(* IEC 61131-3 sources: codesys-api/examples/plc_architecture/bench/st, 5 files *)

(* ---- PRG_BusTask.st ---- *)
PROGRAM PRG_BusTask
// Body of the bus task on the bench (BusTask: cyclic 5 ms, priority between control and comms): PRG_Bus, timed.
// ExecUs is wall time, so it includes time the control task preempted it. Per line: requests and errors per
// second over the last full second, and how long the slowest request took.
VAR
	ResetStats : BOOL;
	ScanCount : UDINT;
	ExecUs : UDINT;
	MaxExecUs : UDINT;
	ExecTotalUs : ULINT;
	MaxIntervalUs : UDINT;
	RequestsPerSecond : ARRAY[1..GVL_Bus.LINE_COUNT] OF UDINT;
	ErrorsPerSecond : ARRAY[1..GVL_Bus.LINE_COUNT] OF UDINT;

	StartUs : ULINT;
	PreviousStartUs : ULINT;
	SecondStartUs : ULINT;
	RequestsAtSecond : ARRAY[1..GVL_Bus.LINE_COUNT] OF UDINT;
	ErrorsAtSecond : ARRAY[1..GVL_Bus.LINE_COUNT] OF UDINT;
	Index : INT;
END_VAR
// ---- implementation ----
StartUs := F_NowUs();
IF ResetStats THEN
	ResetStats := FALSE;
	ScanCount := 0;
	MaxExecUs := 0;
	ExecTotalUs := 0;
	MaxIntervalUs := 0;
	PreviousStartUs := 0;
END_IF
IF PreviousStartUs <> 0 THEN
	MaxIntervalUs := MAX(MaxIntervalUs, ULINT_TO_UDINT(StartUs - PreviousStartUs));
END_IF
PreviousStartUs := StartUs;

PRG_Bus();
PRG_SerialProbe();       // idle unless IsEnabled

IF StartUs - SecondStartUs >= 1000000 THEN
	SecondStartUs := StartUs;
	FOR Index := 1 TO GVL_Bus.LINE_COUNT DO
		RequestsPerSecond[Index] := PRG_Bus.Lines[Index].RequestCount - RequestsAtSecond[Index];
		ErrorsPerSecond[Index] := PRG_Bus.Lines[Index].ErrorCount - ErrorsAtSecond[Index];
		RequestsAtSecond[Index] := PRG_Bus.Lines[Index].RequestCount;
		ErrorsAtSecond[Index] := PRG_Bus.Lines[Index].ErrorCount;
	END_FOR
END_IF

ExecUs := ULINT_TO_UDINT(F_NowUs() - StartUs);
MaxExecUs := MAX(MaxExecUs, ExecUs);
ExecTotalUs := ExecTotalUs + ExecUs;
ScanCount := ScanCount + 1;

(* ---- PRG_CommsTask.st ---- *)
PROGRAM PRG_CommsTask
// Body of the comms task on the two-task bench (CommsTask: cyclic, priority below the control task):
// PRG_Comms, timed. ExecUs is wall time from start to end of this task's scan, so it includes any time the
// control task preempted it. A publish is timed from PRG_Comms.IsRequested going TRUE to FALSE (done).
VAR
	IsEnabled : BOOL := TRUE;
	ResetStats : BOOL;

	ScanCount : UDINT;
	ExecUs : UDINT;
	MaxExecUs : UDINT;
	ExecTotalUs : ULINT;
	MaxIntervalUs : UDINT;
	PublishCount : UDINT;
	LastPublishUs : UDINT;
	MaxPublishUs : UDINT;
	LastPayloadLength : UDINT;
	MaxClientCalls : INT;

	StartUs : ULINT;
	PreviousStartUs : ULINT;
	RequestUs : ULINT;
	WasRequested : BOOL;
END_VAR
// ---- implementation ----
StartUs := F_NowUs();
IF ResetStats THEN
	ResetStats := FALSE;
	ScanCount := 0;
	MaxExecUs := 0;
	ExecTotalUs := 0;
	MaxIntervalUs := 0;
	PublishCount := 0;
	MaxPublishUs := 0;
	MaxClientCalls := 0;
	PreviousStartUs := 0;
END_IF
IF PreviousStartUs <> 0 THEN
	MaxIntervalUs := MAX(MaxIntervalUs, ULINT_TO_UDINT(StartUs - PreviousStartUs));
END_IF
PreviousStartUs := StartUs;

IF IsEnabled THEN
	PRG_Comms();
	MaxClientCalls := MAX(MaxClientCalls, PRG_Comms.ClientCall);
	IF PRG_Comms.IsRequested AND NOT WasRequested THEN
		RequestUs := StartUs;
		LastPayloadLength := PRG_Comms.Used;
	ELSIF WasRequested AND NOT PRG_Comms.IsRequested THEN
		LastPublishUs := ULINT_TO_UDINT(StartUs - RequestUs);
		MaxPublishUs := MAX(MaxPublishUs, LastPublishUs);
		PublishCount := PublishCount + 1;
	END_IF
	WasRequested := PRG_Comms.IsRequested;
END_IF

ExecUs := ULINT_TO_UDINT(F_NowUs() - StartUs);
MaxExecUs := MAX(MaxExecUs, ExecUs);
ExecTotalUs := ExecTotalUs + ExecUs;
ScanCount := ScanCount + 1;

(* ---- PRG_ControlTask.st ---- *)
PROGRAM PRG_ControlTask
// Body of the control task on the two-task bench (MainTask: cyclic 50 ms, priority 1): simulated inputs,
// then the control pipeline, timed. IntervalUs is the start-to-start time of this task; its deviation from
// NominalUs is the jitter the comms task could cause. ExecUs is the time spent in the task.
VAR
	NominalUs : ULINT := 50000;         // the task's configured interval
	ResetStats : BOOL;
	IsQualityCountRequested : BOOL;     // count tags per quality once (costs a pass over the table)

	ScanCount : UDINT;
	IntervalUs : UDINT;
	MinIntervalUs : UDINT := 16#FFFFFFFF;
	MaxIntervalUs : UDINT;
	MaxDeviationUs : UDINT;             // largest |IntervalUs - NominalUs|
	// |IntervalUs - NominalUs| in bands: <= 0.1 ms, 0.5 ms, 1 ms, 2 ms, 5 ms, more
	Deviation : ARRAY[0..5] OF UDINT;
	ExecUs : UDINT;
	MaxExecUs : UDINT;
	ExecTotalUs : ULINT;
	SimUs : UDINT;
	MaxSimUs : UDINT;
	GoodCount : INT;
	NotGoodCount : INT;

	StartUs : ULINT;
	PreviousStartUs : ULINT;
	StepUs : ULINT;
	DeviationUs : UDINT;
	Index : INT;
END_VAR
// ---- implementation ----
StartUs := F_NowUs();
IF ResetStats THEN
	ResetStats := FALSE;
	ScanCount := 0;
	MinIntervalUs := 16#FFFFFFFF;
	MaxIntervalUs := 0;
	MaxDeviationUs := 0;
	FOR Index := 0 TO 5 DO
		Deviation[Index] := 0;
	END_FOR
	MaxExecUs := 0;
	ExecTotalUs := 0;
	MaxSimUs := 0;
	PreviousStartUs := 0;
END_IF
IF PreviousStartUs <> 0 THEN
	IntervalUs := ULINT_TO_UDINT(StartUs - PreviousStartUs);
	MinIntervalUs := MIN(MinIntervalUs, IntervalUs);
	MaxIntervalUs := MAX(MaxIntervalUs, IntervalUs);
	IF UDINT_TO_ULINT(IntervalUs) >= NominalUs THEN
		DeviationUs := IntervalUs - ULINT_TO_UDINT(NominalUs);
	ELSE
		DeviationUs := ULINT_TO_UDINT(NominalUs) - IntervalUs;
	END_IF
	MaxDeviationUs := MAX(MaxDeviationUs, DeviationUs);
	IF DeviationUs <= 100 THEN
		Deviation[0] := Deviation[0] + 1;
	ELSIF DeviationUs <= 500 THEN
		Deviation[1] := Deviation[1] + 1;
	ELSIF DeviationUs <= 1000 THEN
		Deviation[2] := Deviation[2] + 1;
	ELSIF DeviationUs <= 2000 THEN
		Deviation[3] := Deviation[3] + 1;
	ELSIF DeviationUs <= 5000 THEN
		Deviation[4] := Deviation[4] + 1;
	ELSE
		Deviation[5] := Deviation[5] + 1;
	END_IF
END_IF
PreviousStartUs := StartUs;

StepUs := F_NowUs();
PRG_SimInputs();
SimUs := ULINT_TO_UDINT(F_NowUs() - StepUs);
MaxSimUs := MAX(MaxSimUs, SimUs);

PRG_Control();

IF IsQualityCountRequested THEN
	IsQualityCountRequested := FALSE;
	GoodCount := 0;
	NotGoodCount := 0;
	FOR Index := 1 TO GVL_Tags.TAG_COUNT DO
		IF GVL_Tags.Tags[Index].Quality = E_Quality.GOOD THEN
			GoodCount := GoodCount + 1;
		ELSE
			NotGoodCount := NotGoodCount + 1;
		END_IF
	END_FOR
END_IF

ExecUs := ULINT_TO_UDINT(F_NowUs() - StartUs);
MaxExecUs := MAX(MaxExecUs, ExecUs);
ExecTotalUs := ExecTotalUs + ExecUs;
ScanCount := ScanCount + 1;

(* ---- PRG_SerialProbe.st ---- *)
PROGRAM PRG_SerialProbe
// Receive-only check of a PLC serial port, no Modbus: opens the port with SysCom and counts every byte that
// arrives, keeping the last 32. For "the PLC sends but never hears a reply": send a known pattern from the PC
// (bench/serial_pattern.py) and see whether it lands here. Turn the bus line on that port off first
// (PRG_Bus.Lines[n].IsEnabled := FALSE); a port can only be open once. Called from the bus task.
VAR
	IsEnabled : BOOL;                   // set online
	ComPort : INT := 2;
	Baudrate : UDINT := 9600;
	IsVendorSequence : BOOL := TRUE;    // open like AutomationDirect's example (SysComOpen + SysComSetSettings)
	SetResult : UDINT;

	IsOpen : BOOL;
	OpenResult : UDINT;                 // runtime error code of the last open; 0 = OK
	BytesReceived : UDINT;
	ReadCalls : UDINT;
	LastBytes : ARRAY[0..31] OF BYTE;   // most recent bytes, oldest overwritten first
	NextSlot : INT;

	Handle : SysCom.RTS_IEC_HANDLE;
	Settings : SysCom.SysComSettings;
	Result : SysCom.RTS_IEC_RESULT;
	Buffer : ARRAY[0..63] OF BYTE;
	Count : UDINT;
	Index : UDINT;
END_VAR
// ---- implementation ----
IF IsEnabled AND NOT IsOpen THEN
	Settings.sPort := SysCom.SYS_COM_PORTS.SYS_COMPORT1;
	IF ComPort = 2 THEN
		Settings.sPort := SysCom.SYS_COM_PORTS.SYS_COMPORT2;
	END_IF
	Settings.ulBaudrate := SysCom.SYS_COM_BAUDRATE.SYS_BR_9600;
	IF Baudrate = 115200 THEN
		Settings.ulBaudrate := SysCom.SYS_COM_BAUDRATE.SYS_BR_115200;
	END_IF
	Settings.byParity := SysCom.SYS_COM_PARITY.SYS_NOPARITY;
	Settings.byStopBits := SysCom.SYS_COM_STOPBITS.SYS_ONESTOPBIT;
	Settings.ulTimeout := 0;
	Settings.ulBufferSize := 0;
	IF IsVendorSequence THEN
		// AutomationDirect's Demo_SerialPassthrough: open the port, then apply the settings.
		Settings.ulTimeout := 10;
		Handle := SysCom.SysComOpen(sPort := Settings.sPort, pResult := ADR(Result));
		OpenResult := Result;
		IF Result = 0 THEN
			Result := SysCom.SysComSetSettings(hCom := Handle, pSettings := ADR(Settings), pSettingsEx := 0);
			SetResult := Result;
		END_IF
	ELSE
		Handle := SysCom.SysComOpen2(pSettings := ADR(Settings), pSettingsEx := 0, pResult := ADR(Result));
		OpenResult := Result;
	END_IF
	IsOpen := Result = 0;
ELSIF NOT IsEnabled AND IsOpen THEN
	SysCom.SysComClose(hCom := Handle);
	IsOpen := FALSE;
END_IF

IF IsOpen THEN
	Count := SysCom.SysComRead(hCom := Handle, pbyBuffer := ADR(Buffer), ulSize := SIZEOF(Buffer), ulTimeout := 0, pResult := ADR(Result));
	ReadCalls := ReadCalls + 1;
	IF Count > 0 THEN
		FOR Index := 0 TO MIN(Count, SIZEOF(Buffer)) - 1 DO
			LastBytes[NextSlot] := Buffer[Index];
			NextSlot := (NextSlot + 1) MOD 32;
		END_FOR
		BytesReceived := BytesReceived + Count;
	END_IF
END_IF

(* ---- PRG_SimInputs.st ---- *)
PROGRAM PRG_SimInputs
// Bench stand-in for local I/O: the tags of source 0 keep moving. Each scan ChangePerScan of them get a new raw
// value, cycling through the table (100 per 50 ms scan = every tag changes about once a second). Tags of the bus
// devices come from PRG_Bus instead. Values stay inside the generated ranges: BOOL 0/1, INT 0..99,999, REAL raw
// 0..4,999 (scale 0.1 -> 0..499.9).
VAR
	ChangePerScan : INT := 100;
	NextIndex : INT := 1;
	Step : DINT;
	Count : INT;
END_VAR
// ---- implementation ----
Step := Step + 1;
FOR Count := 1 TO ChangePerScan DO
	IF GVL_Tags.TagConfig[NextIndex].Source = 0 THEN
		CASE GVL_Tags.TagConfig[NextIndex].Kind OF
			E_TagKind.BOOL_TAG:
				GVL_Tags.RawInputs[NextIndex] := DINT_TO_REAL((Step + NextIndex) MOD 2);
			E_TagKind.INT_TAG:
				GVL_Tags.RawInputs[NextIndex] := DINT_TO_REAL((Step * 7 + NextIndex) MOD 100000);
		ELSE
			GVL_Tags.RawInputs[NextIndex] := DINT_TO_REAL((Step * 13 + NextIndex * 3) MOD 5000);
		END_CASE
	END_IF
	NextIndex := NextIndex MOD GVL_Tags.TAG_COUNT + 1;
END_FOR
